// TIA Portal V21 export
// export: Created 2026-11-11T00:48:12.6241293Z, ExportSetting WithDefaults, DisplayName Totally Integrated Automation Portal, DisplayVersion V21 Update 3, DisplayName STEP 7 Professional, DisplayVersion V21 Update 3, DisplayName STEP 7 Safety, DisplayVersion V21, DisplayName Tech WebApplication, DisplayVersion V21, DisplayName WinCC Basic/Comfort/Advanced, DisplayVersion V21 Update 3, DisplayName WinCC Unified, DisplayVersion V21 Update 3
FUNCTION_BLOCK "FB_Scl_sl027"   // FB49, SCL
{ S7_Optimized_Access := 'TRUE' }
VERSION : 0.1
// stored: AutoNumber true, IsIECCheckEnabled false, IsRetainMemResEnabled false, MemoryReserve 100, SetENOAutomatically false, UDAEnableTagReadback false
   VAR_INPUT
      v_mn : Time;
      v_in : Time;
      v_mx : Time;
   END_VAR
   VAR_OUTPUT
      v_ret : Time;
   END_VAR
BEGIN
   #v_ret := LIMIT(MN := #v_mn, IN := #v_in, MX := #v_mx);
END_FUNCTION_BLOCK
